INTERFACE I_Compensator EXTENDS I_Module

METHOD M_Calc : ST_PQ			// 목표에 더할 보정량
VAR_INPUT
	i_stView	: ST_GroupView;
END_VAR
END_METHOD

END_INTERFACE

(* stored: Version 1.1.0.1, ProductVersion 3.1.4024.15
   Itf I_Compensator: Id {773f04a9-ad59-43f9-9abd-8e0598413510}
   Method M_Calc: Id {22f575b0-1991-4edb-9b44-5ca76b8fa76d} *)
